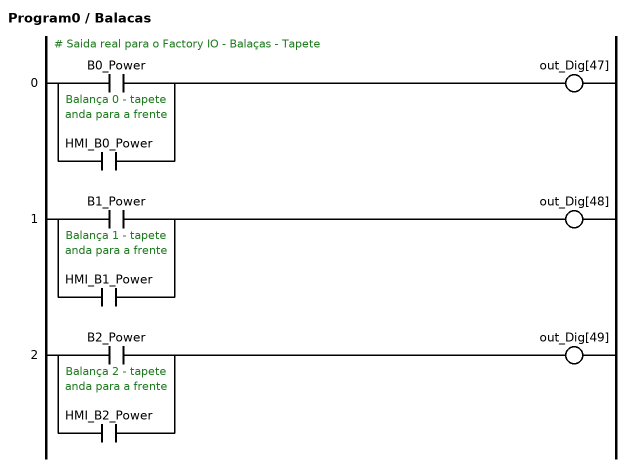
(* [picture p72: Program0 / Balacas, rungs 0-2] *)
(* Rung 0: # Saida real para o Factory IO - Balaças - Tapete *)
out_Dig[47] := B0_Power OR HMI_B0_Power;
(* Rung 1 *)
out_Dig[48] := B1_Power OR HMI_B1_Power;
(* Rung 2 *)
out_Dig[49] := B2_Power OR HMI_B2_Power;

(* Section Laminas_Stop: ladder, written here as Structured Text *)

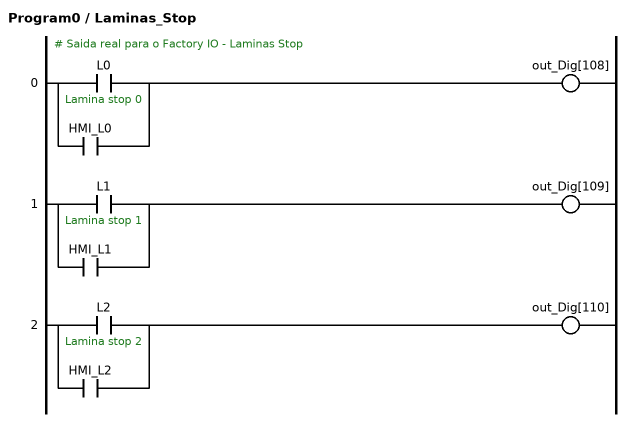
(* Rung 0: # Saida real para o Factory IO - Laminas Stop *)
out_Dig[108] := L0 OR HMI_L0;
(* Rung 1 *)
out_Dig[109] := L1 OR HMI_L1;
(* Rung 2 *)
out_Dig[110] := L2 OR HMI_L2;

(* Section Machines_Centers: ladder, written here as Structured Text *)

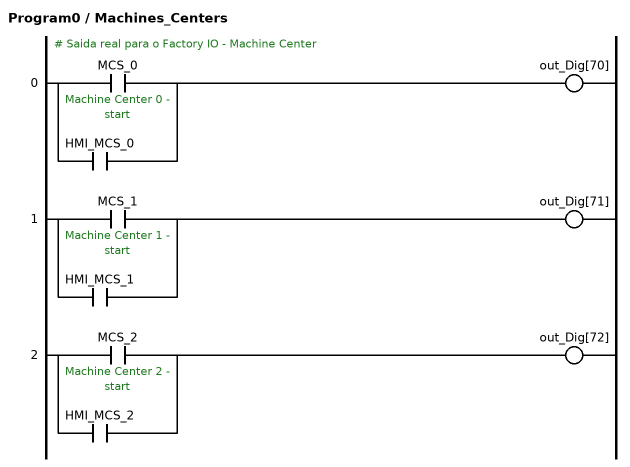
(* Rung 0: # Saida real para o Factory IO - Machine Center *)
out_Dig[70] := MCS_0 OR HMI_MCS_0;
(* Rung 1 *)
out_Dig[71] := MCS_1 OR HMI_MCS_1;
(* Rung 2 *)
out_Dig[72] := MCS_2 OR HMI_MCS_2;

(* Section Arranque_E: ladder, written here as Structured Text *)

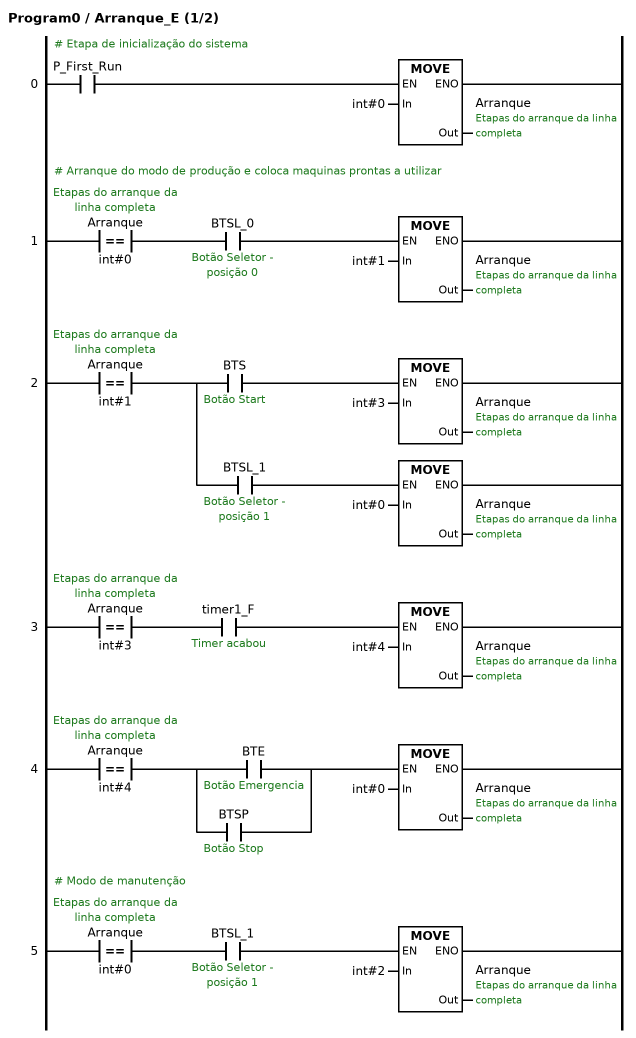
(* Rung 0: # Etapa de inicialização do sistema *)
IF P_First_Run THEN Arranque := int#0; END_IF;
(* Rung 1: # Arranque do modo de produção e coloca maquinas prontas a utilizar *)
IF (Arranque = int#0) AND BTSL_0 THEN Arranque := int#1; END_IF;
(* Rung 2 *)
_p20 := Arranque = int#1;
IF (Arranque = int#1) AND BTS THEN Arranque := int#3; END_IF;
IF _p20 AND BTSL_1 THEN Arranque := int#0; END_IF;
(* Rung 3 *)
IF (Arranque = int#3) AND timer1_F THEN Arranque := int#4; END_IF;
(* Rung 4 *)
IF (Arranque = int#4) AND (BTE OR BTSP) THEN Arranque := int#0; END_IF;
(* Rung 5: # Modo de manutenção *)
IF (Arranque = int#0) AND BTSL_1 THEN Arranque := int#2; END_IF;

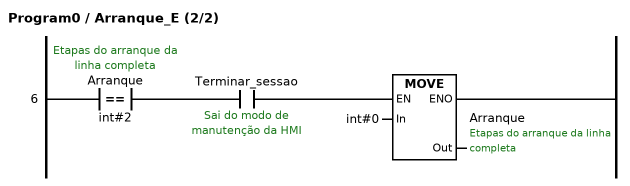
(* Rung 6 *)
IF (Arranque = int#2) AND Terminar_sessao THEN Arranque := int#0; END_IF;

(* Section Arranque_S: ladder, written here as Structured Text *)

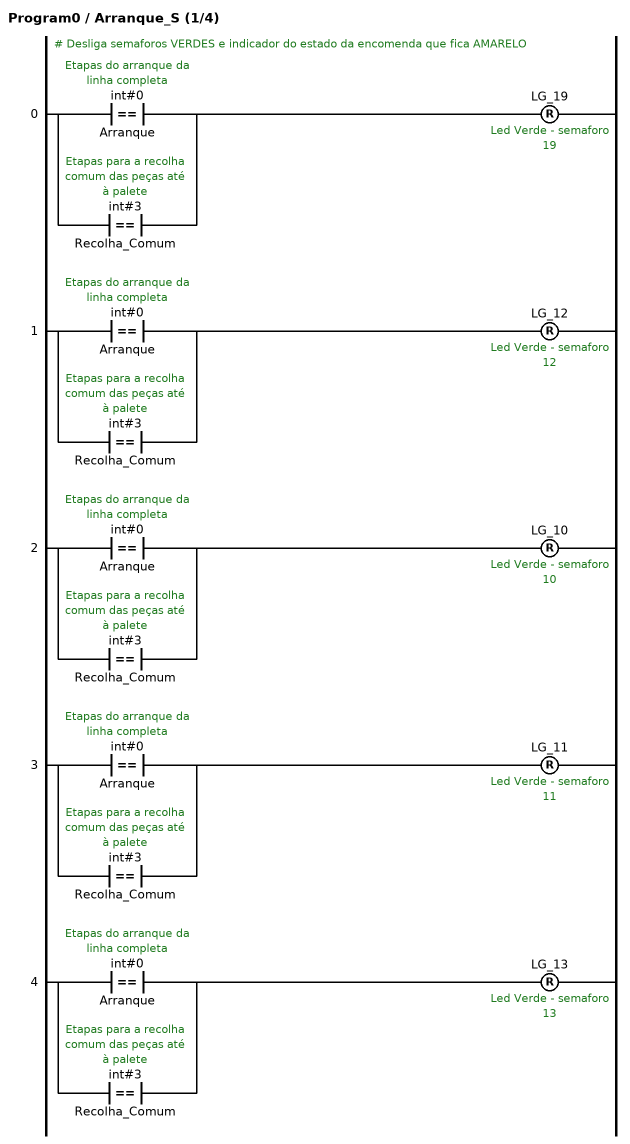
(* Rung 0: # Desliga semaforos VERDES e indicador do estado da encomenda que fica AMARELO *)
IF (int#0 = Arranque) OR (int#3 = Recolha_Comum) THEN LG_19 := FALSE; END_IF;
(* Rung 1 *)
IF (int#0 = Arranque) OR (int#3 = Recolha_Comum) THEN LG_12 := FALSE; END_IF;
(* Rung 2 *)
IF (int#0 = Arranque) OR (int#3 = Recolha_Comum) THEN LG_10 := FALSE; END_IF;
(* Rung 3 *)
IF (int#0 = Arranque) OR (int#3 = Recolha_Comum) THEN LG_11 := FALSE; END_IF;
(* Rung 4 *)
IF (int#0 = Arranque) OR (int#3 = Recolha_Comum) THEN LG_13 := FALSE; END_IF;

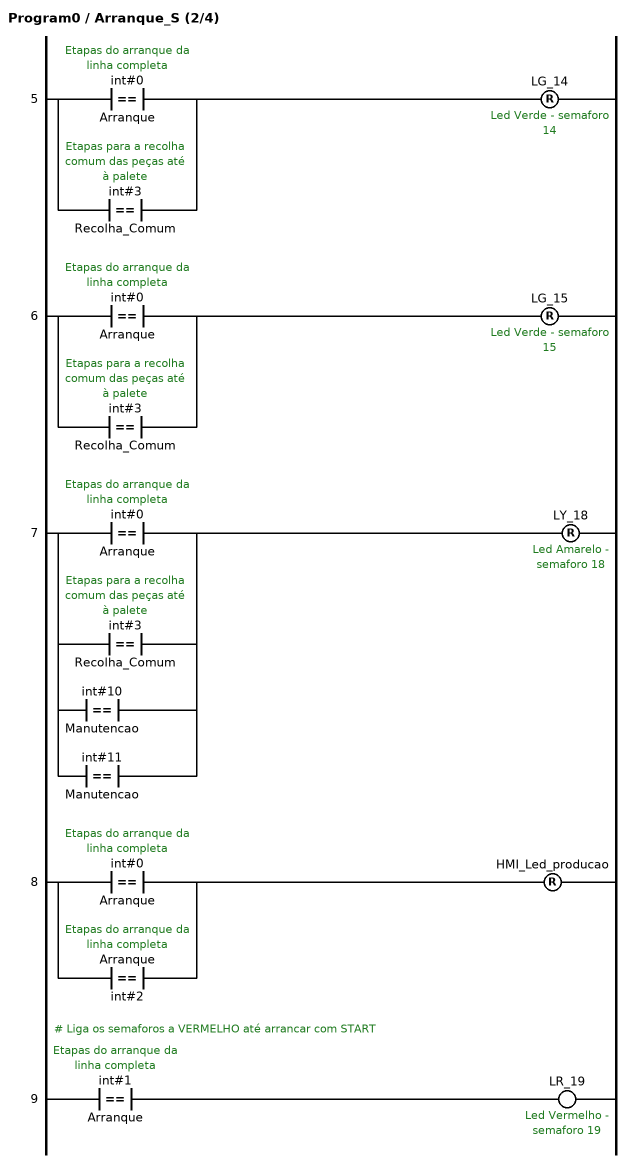
(* Rung 5 *)
IF (int#0 = Arranque) OR (int#3 = Recolha_Comum) THEN LG_14 := FALSE; END_IF;
(* Rung 6 *)
IF (int#0 = Arranque) OR (int#3 = Recolha_Comum) THEN LG_15 := FALSE; END_IF;
(* Rung 7 *)
IF (int#0 = Arranque) OR (int#3 = Recolha_Comum) OR (int#10 = Manutencao) OR (int#11 = Manutencao) THEN
    LY_18 := FALSE;
END_IF;
(* Rung 8 *)
IF (int#0 = Arranque) OR (Arranque = int#2) THEN HMI_Led_producao := FALSE; END_IF;
(* Rung 9: # Liga os semaforos a VERMELHO até arrancar com START *)
LR_19 := int#1 = Arranque;

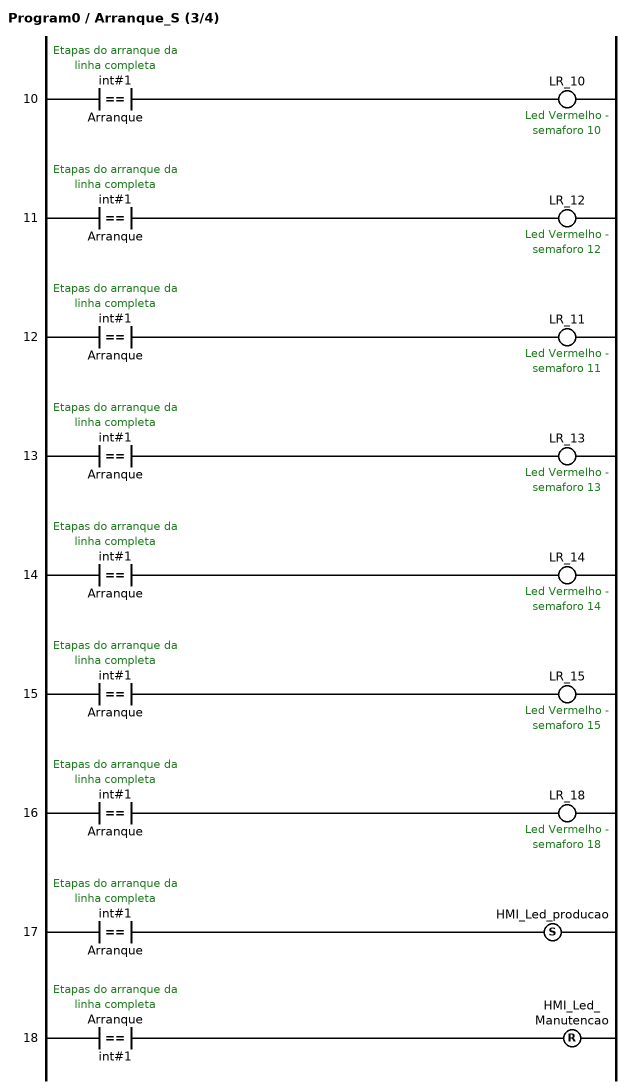
(* Rung 10 *)
LR_10 := int#1 = Arranque;
(* Rung 11 *)
LR_12 := int#1 = Arranque;
(* Rung 12 *)
LR_11 := int#1 = Arranque;
(* Rung 13 *)
LR_13 := int#1 = Arranque;
(* Rung 14 *)
LR_14 := int#1 = Arranque;
(* Rung 15 *)
LR_15 := int#1 = Arranque;
(* Rung 16 *)
LR_18 := int#1 = Arranque;
(* Rung 17 *)
IF int#1 = Arranque THEN HMI_Led_producao := TRUE; END_IF;
(* Rung 18 *)
IF Arranque = int#1 THEN HMI_Led_Manutencao := FALSE; END_IF;

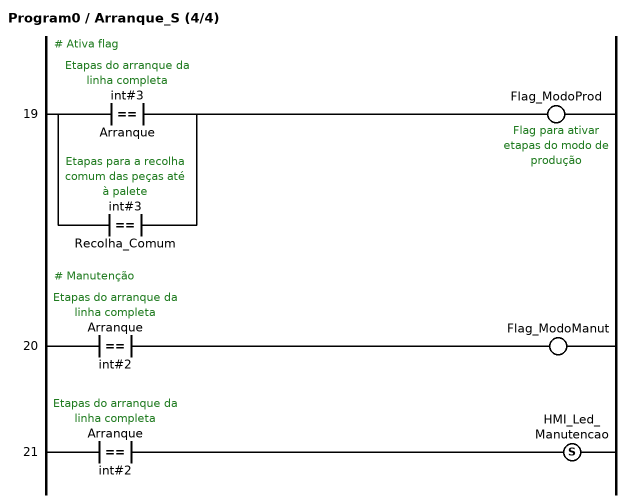
(* Rung 19: # Ativa flag *)
Flag_ModoProd := (int#3 = Arranque) OR (int#3 = Recolha_Comum);
(* Rung 20: # Manutenção *)
Flag_ModoManut := Arranque = int#2;
(* Rung 21 *)
IF Arranque = int#2 THEN HMI_Led_Manutencao := TRUE; END_IF;

(* Section Manutencao_E: ladder, written here as Structured Text *)

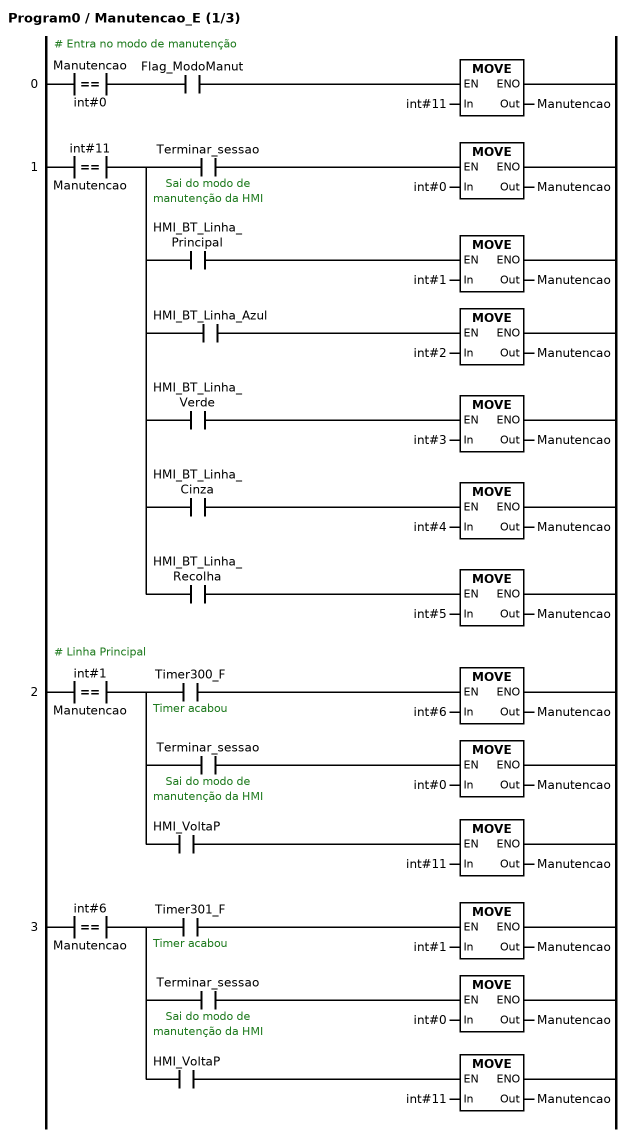
(* Rung 0: # Entra no modo de manutenção *)
IF (Manutencao = int#0) AND Flag_ModoManut THEN Manutencao := int#11; END_IF;
(* Rung 1 *)
_p21 := int#11 = Manutencao;
IF (int#11 = Manutencao) AND Terminar_sessao THEN Manutencao := int#0; END_IF;
IF _p21 AND HMI_BT_Linha_Principal THEN Manutencao := int#1; END_IF;
IF _p21 AND HMI_BT_Linha_Azul THEN Manutencao := int#2; END_IF;
IF _p21 AND HMI_BT_Linha_Verde THEN Manutencao := int#3; END_IF;
IF _p21 AND HMI_BT_Linha_Cinza THEN Manutencao := int#4; END_IF;
IF _p21 AND HMI_BT_Linha_Recolha THEN Manutencao := int#5; END_IF;
(* Rung 2: # Linha Principal *)
_p22 := int#1 = Manutencao;
IF (int#1 = Manutencao) AND Timer300_F THEN Manutencao := int#6; END_IF;
IF _p22 AND Terminar_sessao THEN Manutencao := int#0; END_IF;
IF _p22 AND HMI_VoltaP THEN Manutencao := int#11; END_IF;
(* Rung 3 *)
_p23 := int#6 = Manutencao;
IF (int#6 = Manutencao) AND Timer301_F THEN Manutencao := int#1; END_IF;
IF _p23 AND Terminar_sessao THEN Manutencao := int#0; END_IF;
IF _p23 AND HMI_VoltaP THEN Manutencao := int#11; END_IF;

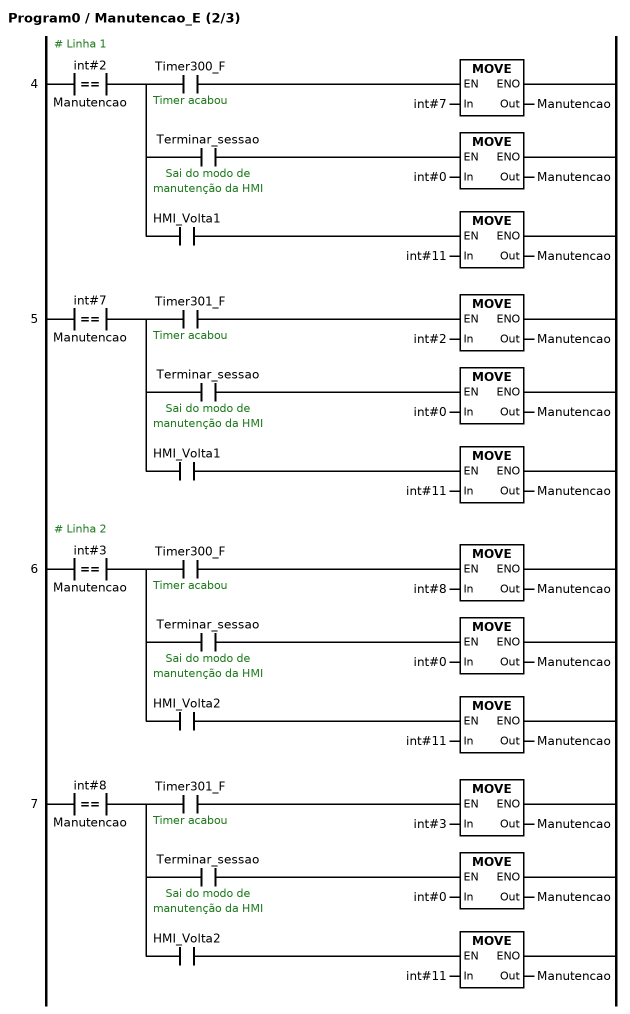
(* Rung 4: # Linha 1 *)
_p24 := int#2 = Manutencao;
IF (int#2 = Manutencao) AND Timer300_F THEN Manutencao := int#7; END_IF;
IF _p24 AND Terminar_sessao THEN Manutencao := int#0; END_IF;
IF _p24 AND HMI_Volta1 THEN Manutencao := int#11; END_IF;
(* Rung 5 *)
_p25 := int#7 = Manutencao;
IF (int#7 = Manutencao) AND Timer301_F THEN Manutencao := int#2; END_IF;
IF _p25 AND Terminar_sessao THEN Manutencao := int#0; END_IF;
IF _p25 AND HMI_Volta1 THEN Manutencao := int#11; END_IF;
(* Rung 6: # Linha 2 *)
_p26 := int#3 = Manutencao;
IF (int#3 = Manutencao) AND Timer300_F THEN Manutencao := int#8; END_IF;
IF _p26 AND Terminar_sessao THEN Manutencao := int#0; END_IF;
IF _p26 AND HMI_Volta2 THEN Manutencao := int#11; END_IF;
(* Rung 7 *)
_p27 := int#8 = Manutencao;
IF (int#8 = Manutencao) AND Timer301_F THEN Manutencao := int#3; END_IF;
IF _p27 AND Terminar_sessao THEN Manutencao := int#0; END_IF;
IF _p27 AND HMI_Volta2 THEN Manutencao := int#11; END_IF;

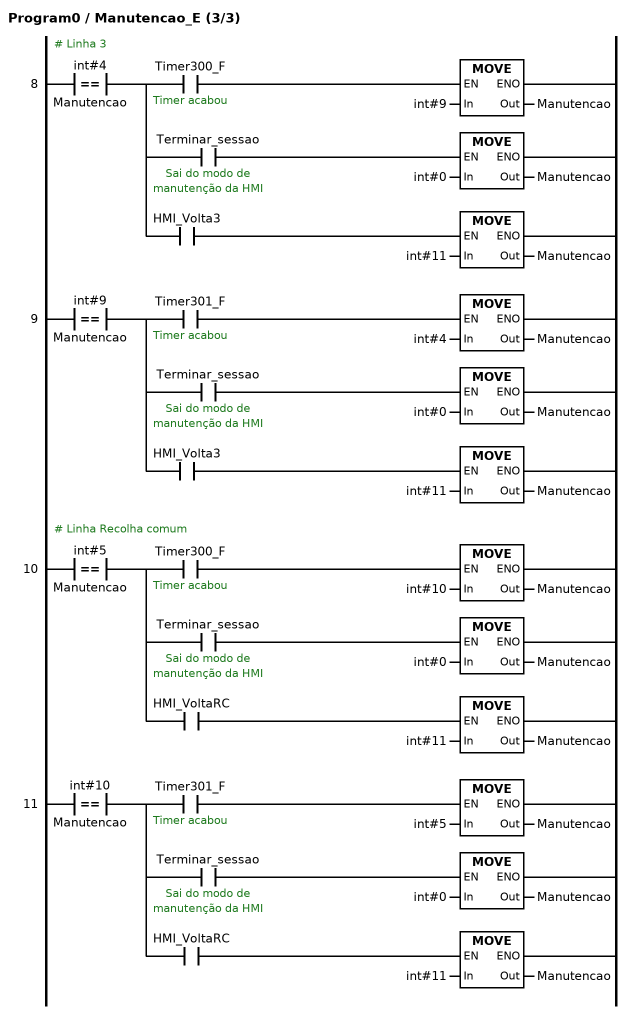
(* Rung 8: # Linha 3 *)
_p28 := int#4 = Manutencao;
IF (int#4 = Manutencao) AND Timer300_F THEN Manutencao := int#9; END_IF;
IF _p28 AND Terminar_sessao THEN Manutencao := int#0; END_IF;
IF _p28 AND HMI_Volta3 THEN Manutencao := int#11; END_IF;
(* Rung 9 *)
_p29 := int#9 = Manutencao;
IF (int#9 = Manutencao) AND Timer301_F THEN Manutencao := int#4; END_IF;
IF _p29 AND Terminar_sessao THEN Manutencao := int#0; END_IF;
IF _p29 AND HMI_Volta3 THEN Manutencao := int#11; END_IF;
(* Rung 10: # Linha Recolha comum *)
_p30 := int#5 = Manutencao;
IF (int#5 = Manutencao) AND Timer300_F THEN Manutencao := int#10; END_IF;
IF _p30 AND Terminar_sessao THEN Manutencao := int#0; END_IF;
IF _p30 AND HMI_VoltaRC THEN Manutencao := int#11; END_IF;
(* Rung 11 *)
_p31 := int#10 = Manutencao;
IF (int#10 = Manutencao) AND Timer301_F THEN Manutencao := int#5; END_IF;
IF _p31 AND Terminar_sessao THEN Manutencao := int#0; END_IF;
IF _p31 AND HMI_VoltaRC THEN Manutencao := int#11; END_IF;

(* Section Tapete_Principal_E: ladder, written here as Structured Text *)

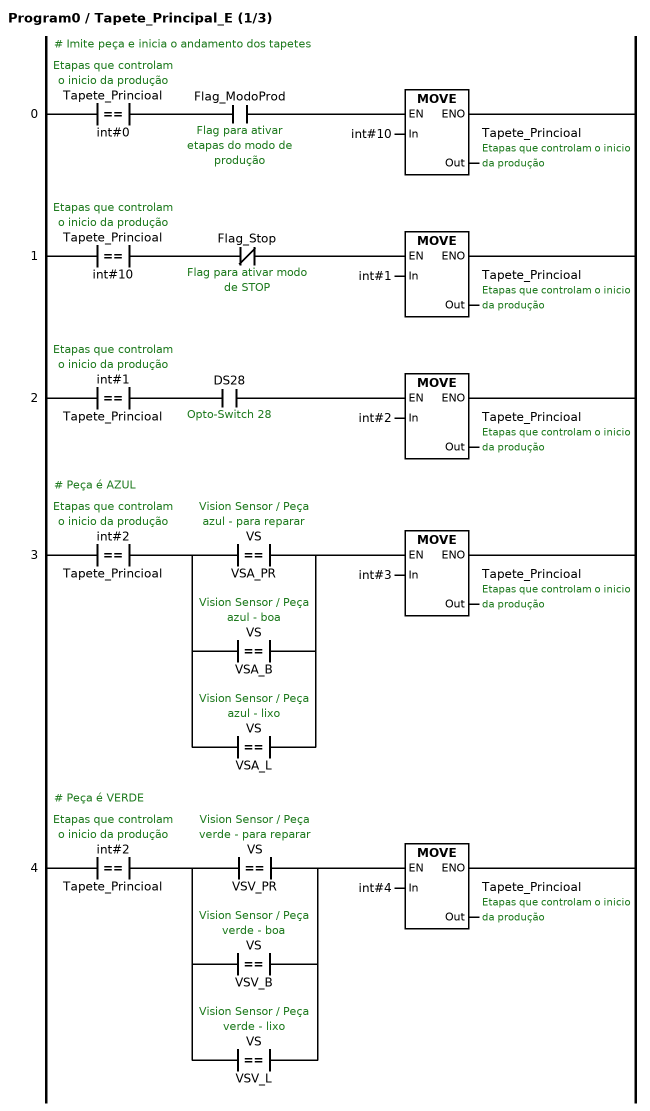
(* Rung 0: # Imite peça e inicia o andamento dos tapetes *)
IF (Tapete_Princioal = int#0) AND Flag_ModoProd THEN Tapete_Princioal := int#10; END_IF;
(* Rung 1 *)
IF (Tapete_Princioal = int#10) AND NOT Flag_Stop THEN Tapete_Princioal := int#1; END_IF;
(* Rung 2 *)
IF (int#1 = Tapete_Princioal) AND DS28 THEN Tapete_Princioal := int#2; END_IF;
(* Rung 3: # Peça é AZUL *)
IF (int#2 = Tapete_Princioal) AND ((VS = VSA_PR) OR (VS = VSA_B) OR (VS = VSA_L)) THEN
    Tapete_Princioal := int#3;
END_IF;
(* Rung 4: # Peça é VERDE *)
IF (int#2 = Tapete_Princioal) AND ((VS = VSV_PR) OR (VS = VSV_B) OR (VS = VSV_L)) THEN
    Tapete_Princioal := int#4;
END_IF;

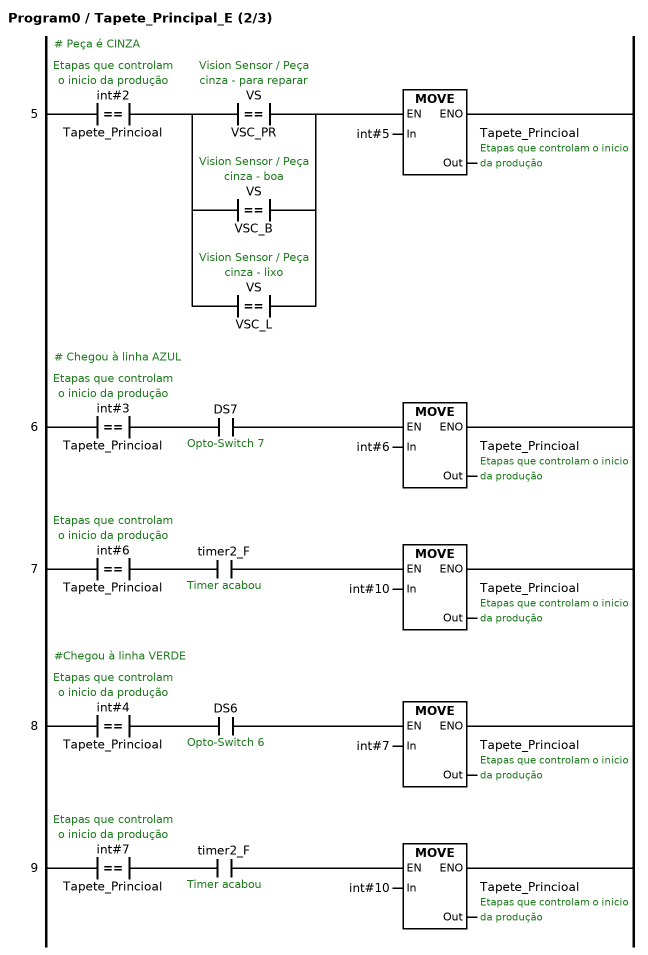
(* Rung 5: # Peça é CINZA *)
IF (int#2 = Tapete_Princioal) AND ((VS = VSC_PR) OR (VS = VSC_B) OR (VS = VSC_L)) THEN
    Tapete_Princioal := int#5;
END_IF;
(* Rung 6: # Chegou à linha AZUL *)
IF (int#3 = Tapete_Princioal) AND DS7 THEN Tapete_Princioal := int#6; END_IF;
(* Rung 7 *)
IF (int#6 = Tapete_Princioal) AND timer2_F THEN Tapete_Princioal := int#10; END_IF;
(* Rung 8: #Chegou à linha VERDE *)
IF (int#4 = Tapete_Princioal) AND DS6 THEN Tapete_Princioal := int#7; END_IF;
(* Rung 9 *)
IF (int#7 = Tapete_Princioal) AND timer2_F THEN Tapete_Princioal := int#10; END_IF;

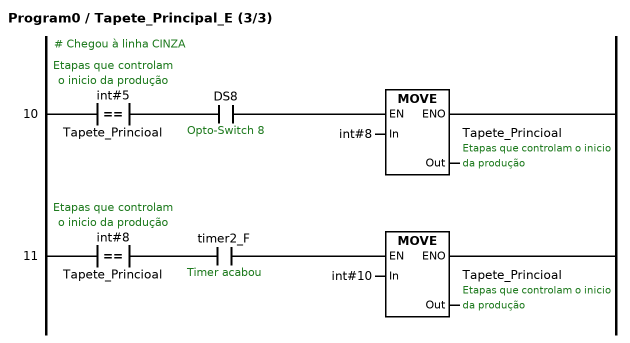
(* Rung 10: # Chegou à linha CINZA *)
IF (int#5 = Tapete_Princioal) AND DS8 THEN Tapete_Princioal := int#8; END_IF;
(* Rung 11 *)
IF (int#8 = Tapete_Princioal) AND timer2_F THEN Tapete_Princioal := int#10; END_IF;

(* Section Tapete_Principal_S: ladder, written here as Structured Text *)

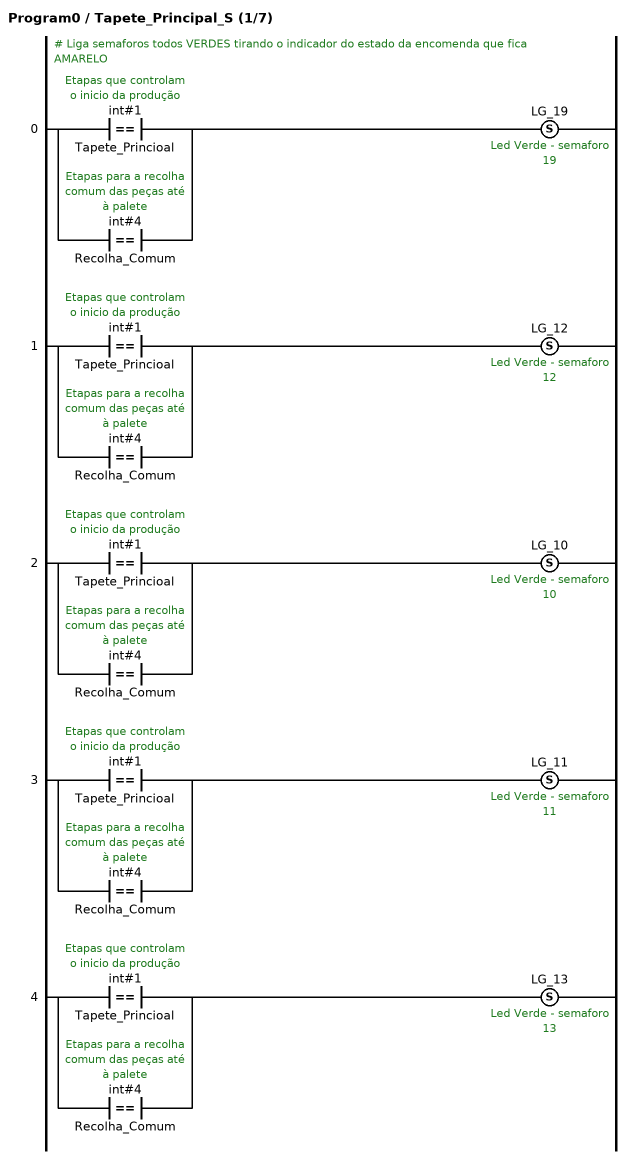
(* Rung 0: # Liga semaforos todos VERDES tirando o indicador do estado da encomenda que fica AMARELO *)
IF (int#1 = Tapete_Princioal) OR (int#4 = Recolha_Comum) THEN LG_19 := TRUE; END_IF;
(* Rung 1 *)
IF (int#1 = Tapete_Princioal) OR (int#4 = Recolha_Comum) THEN LG_12 := TRUE; END_IF;
(* Rung 2 *)
IF (int#1 = Tapete_Princioal) OR (int#4 = Recolha_Comum) THEN LG_10 := TRUE; END_IF;
(* Rung 3 *)
IF (int#1 = Tapete_Princioal) OR (int#4 = Recolha_Comum) THEN LG_11 := TRUE; END_IF;
(* Rung 4 *)
IF (int#1 = Tapete_Princioal) OR (int#4 = Recolha_Comum) THEN LG_13 := TRUE; END_IF;

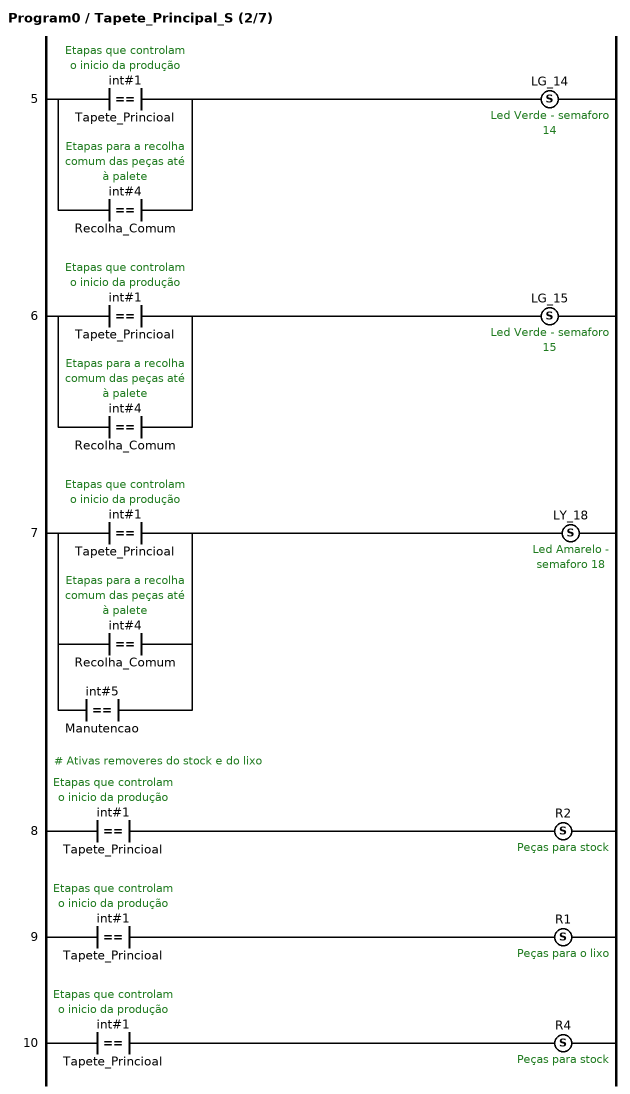
(* Rung 5 *)
IF (int#1 = Tapete_Princioal) OR (int#4 = Recolha_Comum) THEN LG_14 := TRUE; END_IF;
(* Rung 6 *)
IF (int#1 = Tapete_Princioal) OR (int#4 = Recolha_Comum) THEN LG_15 := TRUE; END_IF;
(* Rung 7 *)
IF (int#1 = Tapete_Princioal) OR (int#4 = Recolha_Comum) OR (int#5 = Manutencao) THEN
    LY_18 := TRUE;
END_IF;
(* Rung 8: # Ativas removeres do stock e do lixo *)
IF int#1 = Tapete_Princioal THEN R2 := TRUE; END_IF;
(* Rung 9 *)
IF int#1 = Tapete_Princioal THEN R1 := TRUE; END_IF;
(* Rung 10 *)
IF int#1 = Tapete_Princioal THEN R4 := TRUE; END_IF;

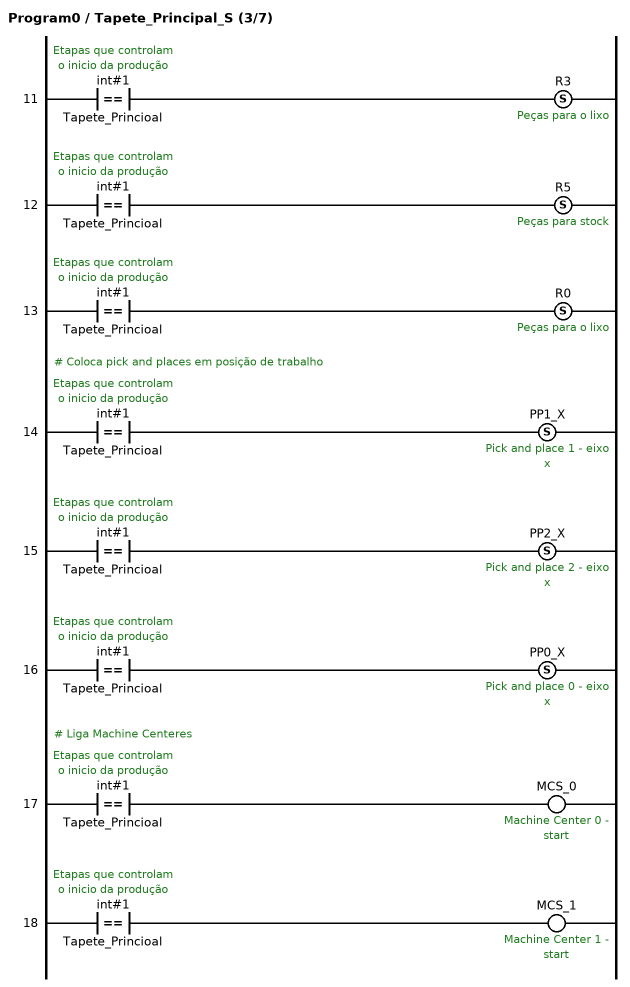
(* Rung 11 *)
IF int#1 = Tapete_Princioal THEN R3 := TRUE; END_IF;
(* Rung 12 *)
IF int#1 = Tapete_Princioal THEN R5 := TRUE; END_IF;
(* Rung 13 *)
IF int#1 = Tapete_Princioal THEN R0 := TRUE; END_IF;
(* Rung 14: # Coloca pick and places em posição de trabalho *)
IF int#1 = Tapete_Princioal THEN PP1_X := TRUE; END_IF;
(* Rung 15 *)
IF int#1 = Tapete_Princioal THEN PP2_X := TRUE; END_IF;
(* Rung 16 *)
IF int#1 = Tapete_Princioal THEN PP0_X := TRUE; END_IF;
(* Rung 17: # Liga Machine Centeres *)
MCS_0 := int#1 = Tapete_Princioal;
(* Rung 18 *)
MCS_1 := int#1 = Tapete_Princioal;

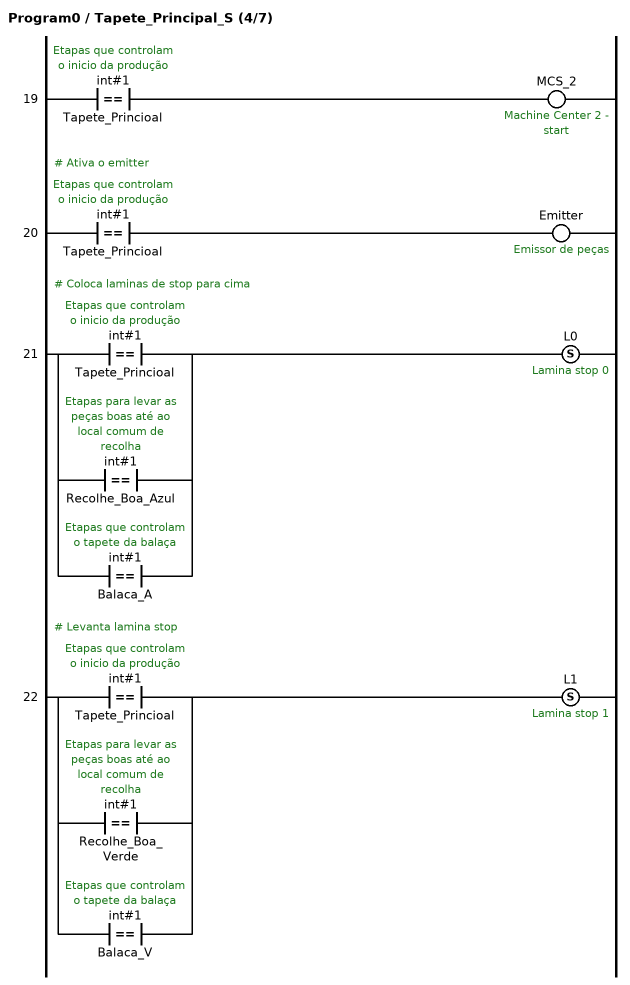
(* Rung 19 *)
MCS_2 := int#1 = Tapete_Princioal;
(* Rung 20: # Ativa o emitter *)
Emitter := int#1 = Tapete_Princioal;
(* Rung 21: # Coloca laminas de stop para cima *)
IF (int#1 = Tapete_Princioal) OR (int#1 = Recolhe_Boa_Azul) OR (int#1 = Balaca_A) THEN L0 := TRUE; END_IF;
(* Rung 22: # Levanta lamina stop *)
IF (int#1 = Tapete_Princioal) OR (int#1 = Recolhe_Boa_Verde) OR (int#1 = Balaca_V) THEN
    L1 := TRUE;
END_IF;

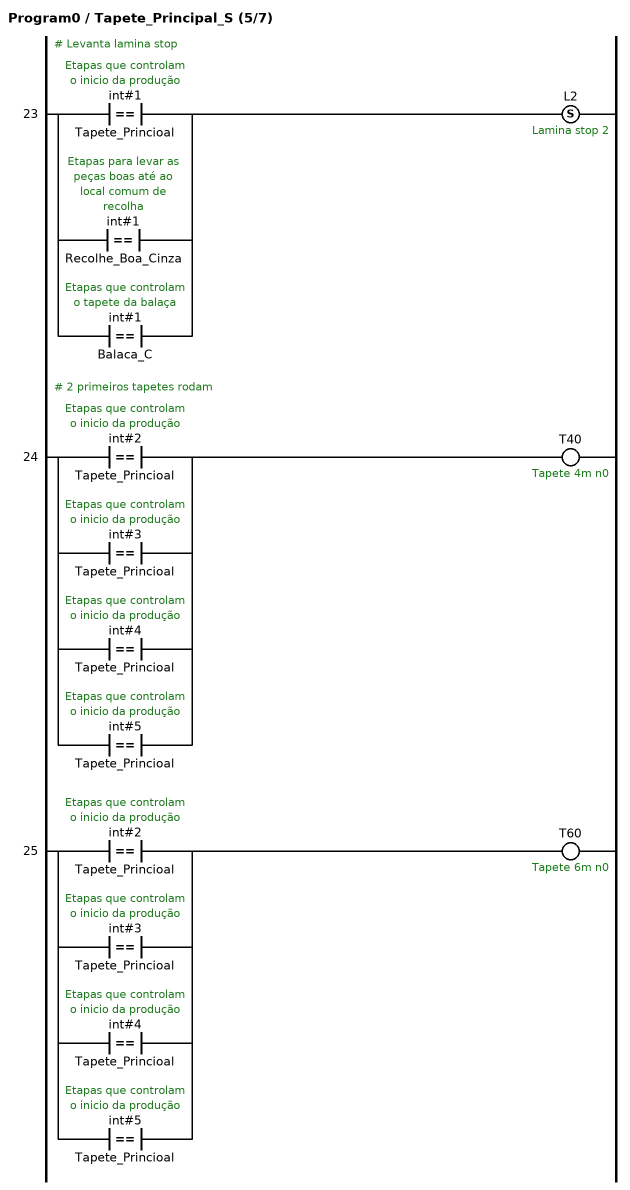
(* Rung 23: # Levanta lamina stop *)
IF (int#1 = Tapete_Princioal) OR (int#1 = Recolhe_Boa_Cinza) OR (int#1 = Balaca_C) THEN
    L2 := TRUE;
END_IF;
(* Rung 24: # 2 primeiros tapetes rodam *)
T40 := (int#2 = Tapete_Princioal) OR (int#3 = Tapete_Princioal) OR (int#4 = Tapete_Princioal) OR (int#5 = Tapete_Princioal);
(* Rung 25 *)
T60 := (int#2 = Tapete_Princioal) OR (int#3 = Tapete_Princioal) OR (int#4 = Tapete_Princioal) OR (int#5 = Tapete_Princioal);

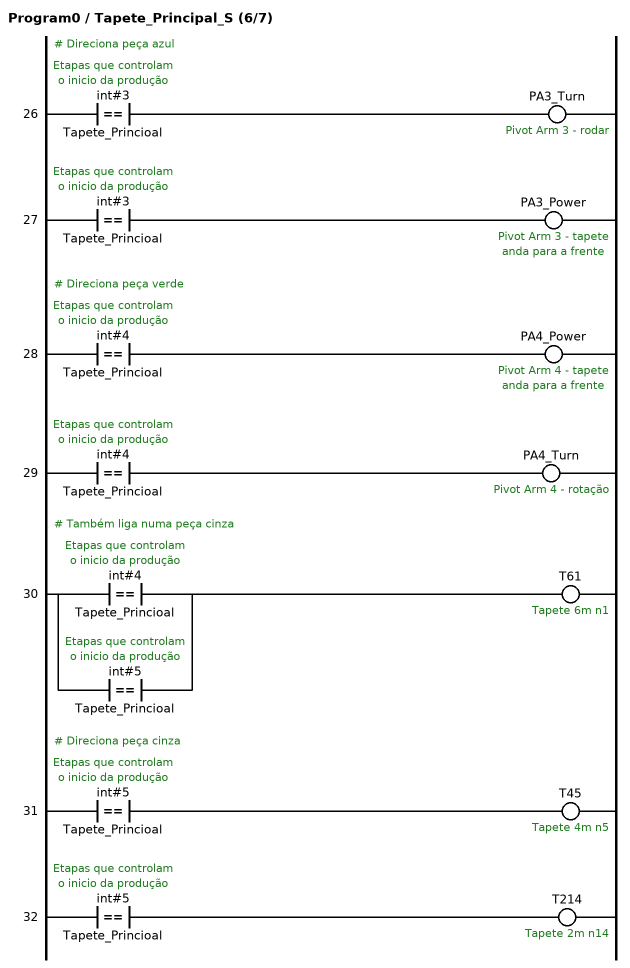
(* Rung 26: # Direciona peça azul *)
PA3_Turn := int#3 = Tapete_Princioal;
(* Rung 27 *)
PA3_Power := int#3 = Tapete_Princioal;
(* Rung 28: # Direciona peça verde *)
PA4_Power := int#4 = Tapete_Princioal;
(* Rung 29 *)
PA4_Turn := int#4 = Tapete_Princioal;
(* Rung 30: # Também liga numa peça cinza *)
T61 := (int#4 = Tapete_Princioal) OR (int#5 = Tapete_Princioal);
(* Rung 31: # Direciona peça cinza *)
T45 := int#5 = Tapete_Princioal;
(* Rung 32 *)
T214 := int#5 = Tapete_Princioal;

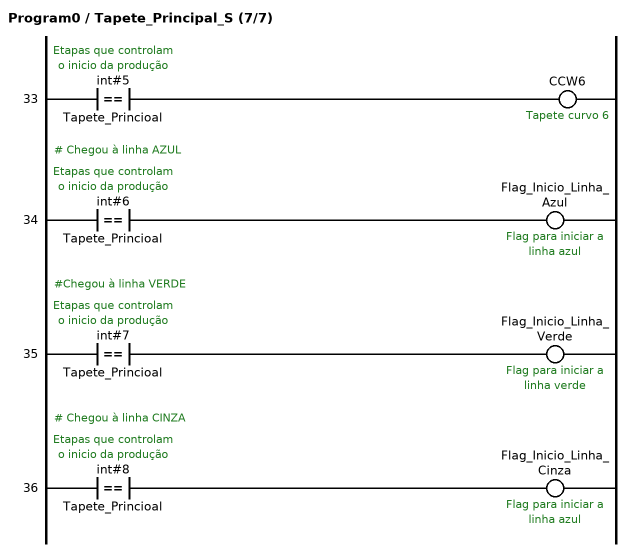
(* Rung 33 *)
CCW6 := int#5 = Tapete_Princioal;
(* Rung 34: # Chegou à linha AZUL *)
Flag_Inicio_Linha_Azul := int#6 = Tapete_Princioal;
(* Rung 35: #Chegou à linha VERDE *)
Flag_Inicio_Linha_Verde := int#7 = Tapete_Princioal;
(* Rung 36: # Chegou à linha CINZA *)
Flag_Inicio_Linha_Cinza := int#8 = Tapete_Princioal;

(* Section Inicio_Linha_E: ladder, written here as Structured Text *)

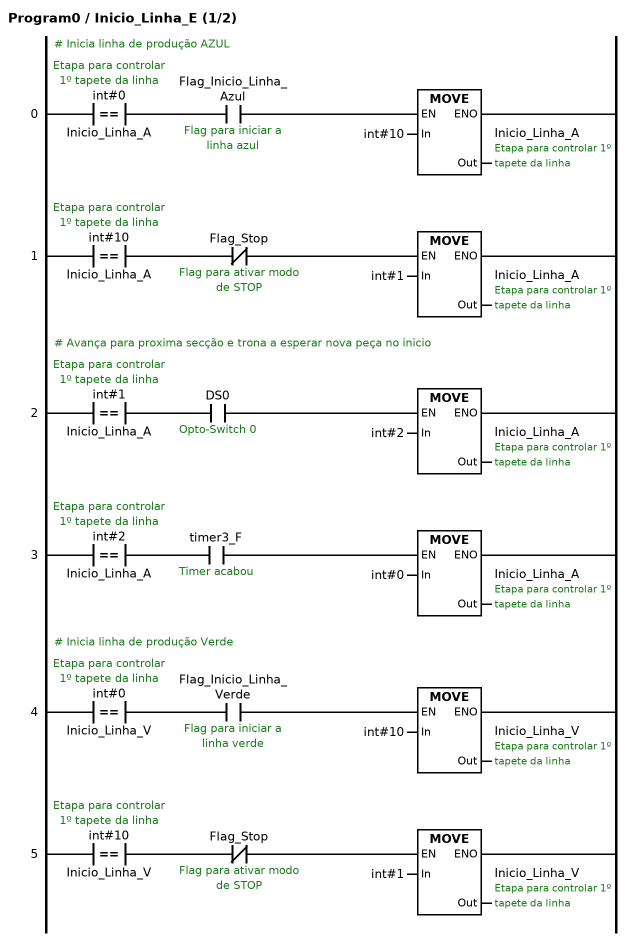
(* Rung 0: # Inicia linha de produção AZUL *)
IF (int#0 = Inicio_Linha_A) AND Flag_Inicio_Linha_Azul THEN Inicio_Linha_A := int#10; END_IF;
(* Rung 1 *)
IF (int#10 = Inicio_Linha_A) AND NOT Flag_Stop THEN Inicio_Linha_A := int#1; END_IF;
(* Rung 2: # Avança para proxima secção e trona a esperar nova peça no inicio *)
IF (int#1 = Inicio_Linha_A) AND DS0 THEN Inicio_Linha_A := int#2; END_IF;
(* Rung 3 *)
IF (int#2 = Inicio_Linha_A) AND timer3_F THEN Inicio_Linha_A := int#0; END_IF;
(* Rung 4: # Inicia linha de produção Verde *)
IF (int#0 = Inicio_Linha_V) AND Flag_Inicio_Linha_Verde THEN Inicio_Linha_V := int#10; END_IF;
(* Rung 5 *)
IF (int#10 = Inicio_Linha_V) AND NOT Flag_Stop THEN Inicio_Linha_V := int#1; END_IF;

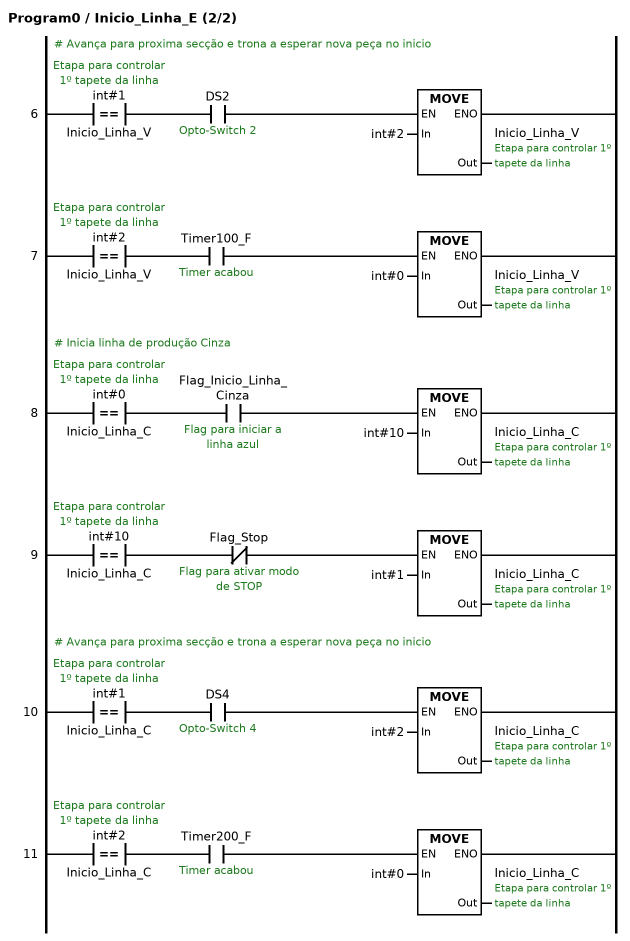
(* Rung 6: # Avança para proxima secção e trona a esperar nova peça no inicio *)
IF (int#1 = Inicio_Linha_V) AND DS2 THEN Inicio_Linha_V := int#2; END_IF;
(* Rung 7 *)
IF (int#2 = Inicio_Linha_V) AND Timer100_F THEN Inicio_Linha_V := int#0; END_IF;
(* Rung 8: # Inicia linha de produção Cinza *)
IF (int#0 = Inicio_Linha_C) AND Flag_Inicio_Linha_Cinza THEN Inicio_Linha_C := int#10; END_IF;
(* Rung 9 *)
IF (int#10 = Inicio_Linha_C) AND NOT Flag_Stop THEN Inicio_Linha_C := int#1; END_IF;
(* Rung 10: # Avança para proxima secção e trona a esperar nova peça no inicio *)
IF (int#1 = Inicio_Linha_C) AND DS4 THEN Inicio_Linha_C := int#2; END_IF;
(* Rung 11 *)
IF (int#2 = Inicio_Linha_C) AND Timer200_F THEN Inicio_Linha_C := int#0; END_IF;

(* Section Inicio_Linha_S: ladder, written here as Structured Text *)

